// TIA Portal V16 export
// export: Created 2000-01-01T00:00:00.0000000Z, ExportSetting None
FUNCTION "FC_Rung" : Void   // FC42, LAD
{ S7_Optimized_Access := 'TRUE' }
   VAR_INPUT
      Local : Int;
   END_VAR
BEGIN

REGION Network 1
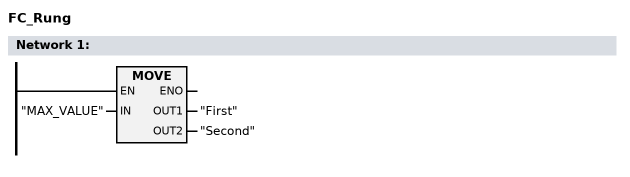
   RUNG wire#powerrail
      Move(in := "MAX_VALUE", out1 => "First", out2 => "Second")
   END_RUNG
   // the same network as SCL:
   "First" := "MAX_VALUE";
   "Second" := "MAX_VALUE";
END_REGION
END_FUNCTION
